// TIA Portal V20 export
// export: Created 2026-10-12T05:11:19.3289455Z, ExportSetting WithDefaults, DisplayName Totally Integrated Automation Portal, DisplayVersion V20, DisplayName TIA Portal Openness, DisplayVersion V20, DisplayName TIA Portal Teamcenter Gateway, DisplayVersion V20, DisplayName TIA Portal Version Control Interface, DisplayVersion V20, DisplayName SINAMICS Startdrive Advanced, DisplayVersion V20 SP1 Update 2, DisplayName SINAMICS Startdrive G110M, G120, G120C, G120D, G120P, G115D, DisplayVersion V20 SP1 Update 2, DisplayName SINAMICS Startdrive G130, G150, S120, S150, SINAMICS MV, G220, S200, S210, DisplayVersion V20 SP1 Update 2, DisplayName STEP 7 Professional, DisplayVersion V20, DisplayName STEP 7 Safety, DisplayVersion V20, DisplayName WinCC Basic/Comfort/Advanced, DisplayVersion V20, DisplayName WinCC Professional, DisplayVersion V20, DisplayName WinCC Unified, DisplayVersion V20
FUNCTION "FRK_State" : Bool   // FC22, SCL
{ S7_Optimized_Access := 'TRUE' }
VERSION : 0.1
// stored: AutoNumber true, IsIECCheckEnabled false, SetENOAutomatically false, UDAEnableTagReadback false
   VAR_INPUT
      Idx : Int;
      Key : String;
      Ok : Bool;
   END_VAR
   VAR_IN_OUT
      Flags : Array[1..12] of "ST_StateFlag";
      Count : Int;
      Touched : Array[1..12] of Bool;
   END_VAR
   VAR_TEMP
      Stamp : DTL;
      ResultCode : Int;
   END_VAR
BEGIN

   #FRK_State := #Ok;
   IF #Idx < 1 OR #Idx > 12 OR LEN(#Key) = 0 OR LEN(#Key) > 120 THEN
       RETURN;
   END_IF;
   IF #Idx > #Count THEN
       #Count := #Idx;
   END_IF;
   IF #Flags[#Idx].Value <> #Ok OR #Flags[#Idx].Key <> #Key OR #Flags[#Idx].Stale THEN
       #Flags[#Idx].Since := LDT#1970-01-01-00:00:00.000000000;
       #ResultCode := RD_SYS_T(OUT => #Stamp);
       IF #ResultCode = 0 THEN
           #Flags[#Idx].Since := DTL_TO_LDT(#Stamp);
       END_IF;
   END_IF;
   #Flags[#Idx].Key := #Key;
   #Flags[#Idx].Value := #Ok;
   #Flags[#Idx].Stale := FALSE;
   #Touched[#Idx] := TRUE;
END_FUNCTION
